Fanuc KAREL source: kt00751.KL

-- PROVISIONAL review KL for V940-1; original PC SHA256 f9b136733fad0e9ee6cd13cf5b1feca862e48c1878712abb99d19aab7fe7fb8d
-- Incomplete behavior may be omitted. Consult companion uncertainty JSON. Do not deploy.
PROGRAM KT00751
%NOLOCKGROUP
VAR
  R1 : REAL
  R2 : REAL
  OUT : REAL
BEGIN
  -- V9_ZERO_TABLE_METADATA_HINT layout=0001; no indexed target words; source/name/runtime held
  -- UNRESOLVED_PC offsets 5-16; opcodes 2E,23
  -- UNRESOLVED_PC offsets 21-32; opcodes 2E,23
  -- UNRESOLVED_PC offsets 37-48; opcodes 2E,23
  -- UNRESOLVED_PC offsets 53-64; opcodes 2E,23
  -- UNRESOLVED_PC offsets 69-82; opcodes 21,67,23
  -- UNRESOLVED_PC offsets 87-91; opcodes 7F
END KT00751
